// TIA Portal V20 export
FUNCTION_BLOCK "PR_LoadingSeq_Soft2.0 1_workflow_95d36b"   // FB48, LAD
{ S7_Optimized_Access := 'TRUE' }
// stored: MemoryReserve 100, SetENOAutomatically false
   VAR_INPUT
      iAbort : Bool;
      iAcceptPartPresent : Bool;
      iAutoRunning : Bool;
      iFaultReset : Bool;
      iLoadGantrySafe : Bool;
      iOTS_Frm_Prev : Bool;
      iPartPresent : Bool;
      iPartPresentInGrip : Bool;
      iRFWriteDone : Bool;
      iRFWriteError : Bool;
      iReject : Bool;
      iReset_fault : Bool;
      iRetry : Bool;
      iRetryCount : Int;
      iSstMode : Bool;
      iSstPB : Bool;
      iStartFrmFibroseq : Bool;
   END_VAR
   VAR_OUTPUT
      qError : Array[0..1] of Bool;
      qLoadingOver : Bool;
      qMessage : Array[0..1] of Bool;
      qRTR_To_Prev : Bool;
   END_VAR
   VAR
      c121_WaitForRFIDWriteOver_T1 : Bool;
      c121_WaitForRFIDWriteOver_T2 : Bool;
      c122_CheckRetryCountOver_T1 : Bool;
      c122_CheckRetryCountOver_T2 : Bool;
      c123_WaitForOperatorDecision_T1 : Bool;
      c123_WaitForOperatorDecision_T2 : Bool;
      c20_CheckRecoveryStatus_T1 : Bool;
      c20_CheckRecoveryStatus_T2 : Bool;
      c20_CheckRecoveryStatus_T3 : Bool;
      c50_CheckPartPresentAtStation_T1 : Bool;
      c50_CheckPartPresentAtStation_T2 : Bool;
      c90_ConfirmPartLoad_T1 : Bool;
      c90_ConfirmPartLoad_T2 : Bool;
      StateNo : Int;
      s100_WaitForOperatorDecision : Bool;
      s100_WaitForOperatorDecision_T1 : Bool;
      s100_WaitForOperatorDecision_T2 : Bool;
      s10_WaitForStartFrmFibroMainSeq : Bool;
      s10_WaitForStartFrmFibroMainSeq_T1 : Bool;
      s120_WaitForGantrySafe : Bool;
      s120_WaitForGantrySafe_T1 : Bool;
      s121_WaitForRFIDWriteOver : Bool;
      s121_WaitForRFIDWriteOver_T1 : Bool;
      s121_WaitForRFIDWriteOver_T2 : Bool;
      s122_CheckRetryCountOver : Bool;
      s122_CheckRetryCountOver_T1 : Bool;
      s122_CheckRetryCountOver_T2 : Bool;
      s123_WaitForOperatorDecision : Bool;
      s123_WaitForOperatorDecision_T1 : Bool;
      s123_WaitForOperatorDecision_T2 : Bool;
      s130_WaitForStartLow : Bool;
      s130_WaitForStartLow_T1 : Bool;
      s1_WaitForResetRelease : Bool;
      s1_WaitForResetRelease_T1 : Bool;
      s20_CheckRecoveryStatus : Bool;
      s20_CheckRecoveryStatus_T1 : Bool;
      s20_CheckRecoveryStatus_T2 : Bool;
      s20_CheckRecoveryStatus_T3 : Bool;
      s30_WaitForOperatorAck : Bool;
      s30_WaitForOperatorAck_T1 : Bool;
      s40_WaitForLoadingGantrySafe : Bool;
      s40_WaitForLoadingGantrySafe_T1 : Bool;
      s50_CheckPartPresentAtStation : Bool;
      s50_CheckPartPresentAtStation_T1 : Bool;
      s50_CheckPartPresentAtStation_T2 : Bool;
      s60_WaitForPartAbsentAndAck : Bool;
      s60_WaitForPartAbsentAndAck_T1 : Bool;
      s70_WaitForOTSFromGantry : Bool;
      s70_WaitForOTSFromGantry_T1 : Bool;
      s80_WaitForPartLoad : Bool;
      s80_WaitForPartLoad_T1 : Bool;
      s90_ConfirmPartLoad : Bool;
      s90_ConfirmPartLoad_T1 : Bool;
      s90_ConfirmPartLoad_T2 : Bool;
      sAbnormalStatus : Bool;
      sLoadInProgress : Bool;
      sLoadInProgressInternal : Int;
      sPartPresent : Bool;
      sRFWriteRetryCount : Int;
      sSst : Bool;
      sSstPulse : Bool;
      sSstRise : Bool;
      sStWtResetRel : Bool;
      sStWtResetRel_T1 : Bool;
   END_VAR
   VAR_TEMP
      tOne : Bool;
   END_VAR
   VAR_TEMP   // added for the SCL form of the ladder/FBD networks
      _w1 : Bool;
      _w2 : Bool;
   END_VAR
BEGIN

REGION Network 1
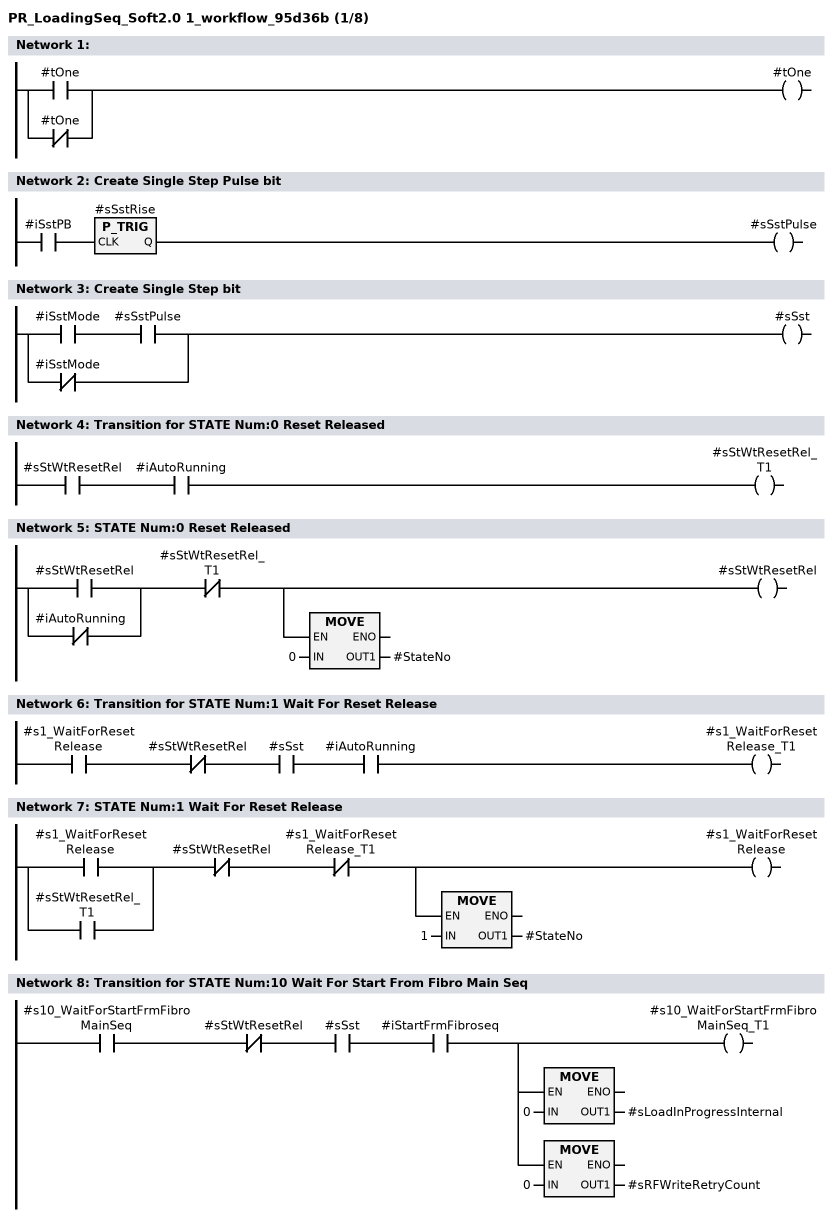
   RUNG wire#powerrail
      Contact( #tOne )
      wire#w1
      Coil( #tOne )
   END_RUNG
   RUNG wire#powerrail
      I_Contact( #tOne )
   END_RUNG wire#w1
   // the same network as SCL:
   #tOne := #tOne OR NOT #tOne;
END_REGION

REGION Network 2: Create Single Step Pulse bit
   RUNG wire#powerrail
      Contact( #iSstPB )
      P_Trig( #sSstRise )
      Coil( #sSstPulse )
   END_RUNG
   // the same network as SCL:
   #_w1 := #iSstPB AND NOT #sSstRise;   // rising edge
   #sSstRise := #iSstPB;
   #sSstPulse := #_w1;
END_REGION

REGION Network 3: Create Single Step bit
   RUNG wire#powerrail
      Contact( #iSstMode )
      Contact( #sSstPulse )
      wire#w1
      Coil( #sSst )
   END_RUNG
   RUNG wire#powerrail
      I_Contact( #iSstMode )
   END_RUNG wire#w1
   // the same network as SCL:
   #sSst := (#iSstMode AND #sSstPulse) OR NOT #iSstMode;
END_REGION

REGION Network 4: Transition for STATE Num:0 Reset Released
   RUNG wire#powerrail
      Contact( #sStWtResetRel )
      Contact( #iAutoRunning )
      Coil( #sStWtResetRel_T1 )
   END_RUNG
   // the same network as SCL:
   #sStWtResetRel_T1 := #sStWtResetRel AND #iAutoRunning;
END_REGION

REGION Network 5: STATE Num:0 Reset Released
   RUNG wire#powerrail
      Contact( #sStWtResetRel )
      wire#w1
      I_Contact( #sStWtResetRel_T1 )
      wire#w2
      Coil( #sStWtResetRel )
   END_RUNG
   RUNG wire#powerrail
      I_Contact( #iAutoRunning )
   END_RUNG wire#w1
   RUNG wire#w2
      { S7_GenerateENO := "TRUE" } Move(in := 0, out1 => #StateNo)
   END_RUNG
   // the same network as SCL:
   #sStWtResetRel := (#sStWtResetRel OR NOT #iAutoRunning) AND NOT #sStWtResetRel_T1;
   IF #sStWtResetRel THEN #StateNo := 0; END_IF;
END_REGION

REGION Network 6: Transition for STATE Num:1 Wait For Reset Release
   RUNG wire#powerrail
      Contact( #s1_WaitForResetRelease )
      I_Contact( #sStWtResetRel )
      Contact( #sSst )
      Contact( #iAutoRunning )
      Coil( #s1_WaitForResetRelease_T1 )
   END_RUNG
   // the same network as SCL:
   #s1_WaitForResetRelease_T1 := #s1_WaitForResetRelease AND NOT #sStWtResetRel AND #sSst AND #iAutoRunning;
END_REGION

REGION Network 7: STATE Num:1 Wait For Reset Release
   RUNG wire#powerrail
      Contact( #s1_WaitForResetRelease )
      wire#w1
      I_Contact( #sStWtResetRel )
      I_Contact( #s1_WaitForResetRelease_T1 )
      wire#w2
      Coil( #s1_WaitForResetRelease )
   END_RUNG
   RUNG wire#powerrail
      Contact( #sStWtResetRel_T1 )
   END_RUNG wire#w1
   RUNG wire#w2
      { S7_GenerateENO := "TRUE" } Move(in := 1, out1 => #StateNo)
   END_RUNG
   // the same network as SCL:
   #s1_WaitForResetRelease := (#s1_WaitForResetRelease OR #sStWtResetRel_T1) AND NOT #sStWtResetRel AND NOT #s1_WaitForResetRelease_T1;
   IF #s1_WaitForResetRelease THEN #StateNo := 1; END_IF;
END_REGION

REGION Network 8: Transition for STATE Num:10 Wait For Start From Fibro Main Seq
   RUNG wire#powerrail
      Contact( #s10_WaitForStartFrmFibroMainSeq )
      I_Contact( #sStWtResetRel )
      Contact( #sSst )
      Contact( #iStartFrmFibroseq )
      wire#w1
      Coil( #s10_WaitForStartFrmFibroMainSeq_T1 )
   END_RUNG
   RUNG wire#w1
      Move(in := 0, out1 => #sLoadInProgressInternal)
   END_RUNG
   RUNG wire#w1
      Move(in := 0, out1 => #sRFWriteRetryCount)
   END_RUNG
   // the same network as SCL:
   #s10_WaitForStartFrmFibroMainSeq_T1 := #s10_WaitForStartFrmFibroMainSeq AND NOT #sStWtResetRel AND #sSst AND #iStartFrmFibroseq;
   IF #s10_WaitForStartFrmFibroMainSeq_T1 THEN
       #sLoadInProgressInternal := 0;
       #sRFWriteRetryCount := 0;
   END_IF;
END_REGION

REGION Network 9: STATE Num:10 Wait For Start From Fibro Main Seq
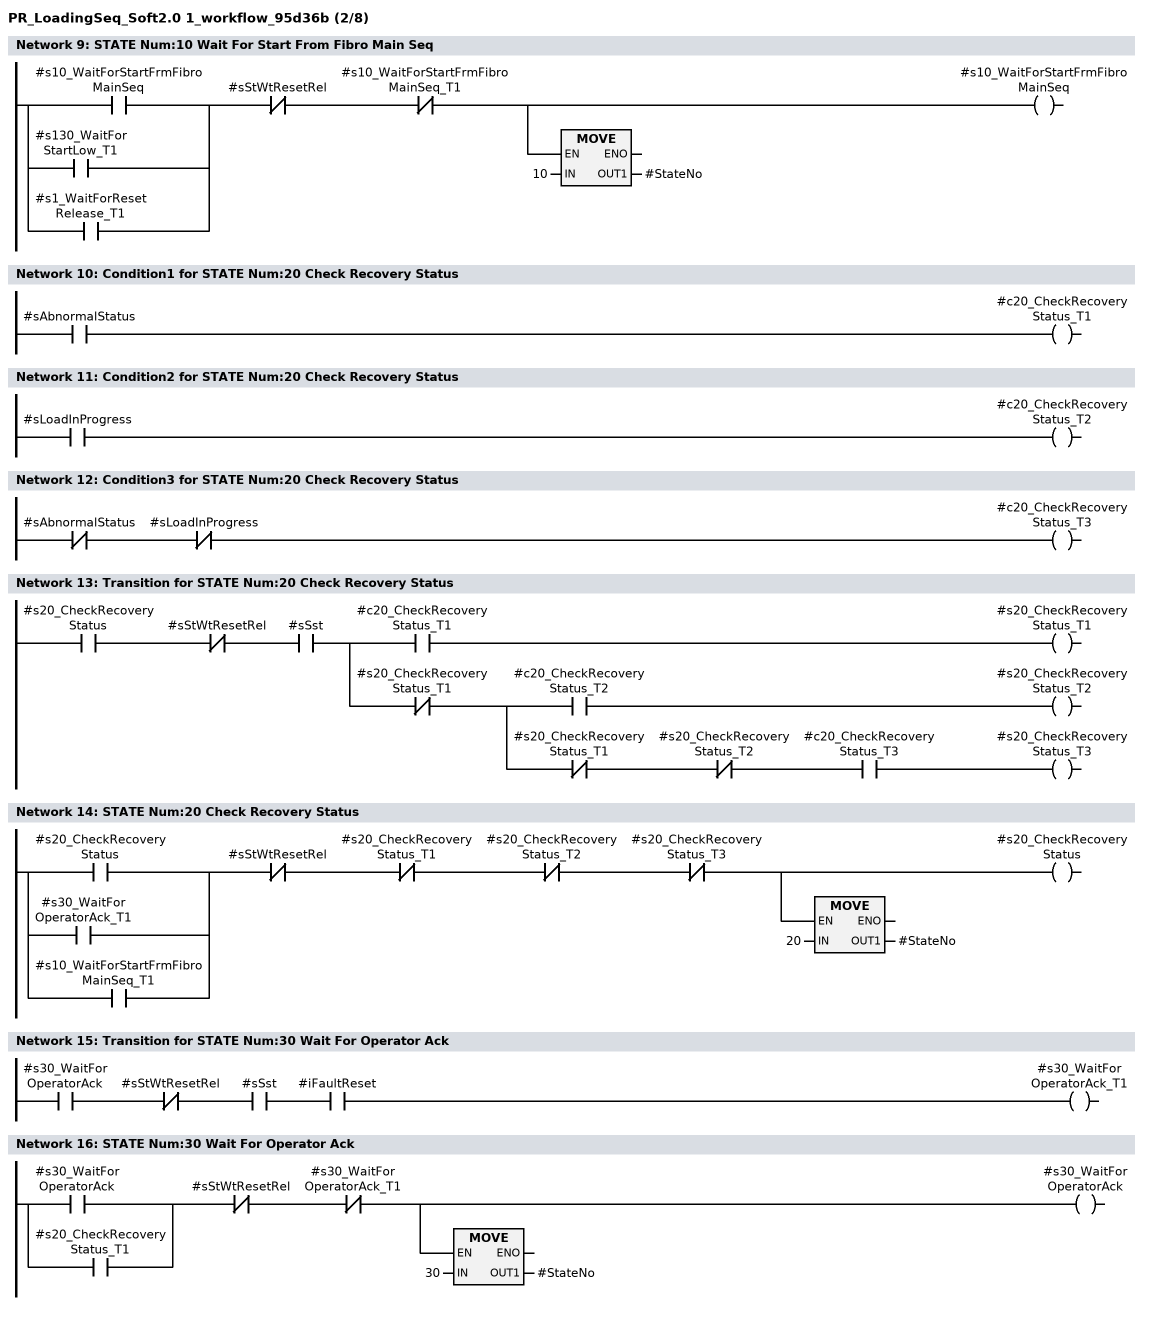
   RUNG wire#powerrail
      Contact( #s10_WaitForStartFrmFibroMainSeq )
      wire#w1
      I_Contact( #sStWtResetRel )
      I_Contact( #s10_WaitForStartFrmFibroMainSeq_T1 )
      wire#w2
      Coil( #s10_WaitForStartFrmFibroMainSeq )
   END_RUNG
   RUNG wire#powerrail
      Contact( #s130_WaitForStartLow_T1 )
   END_RUNG wire#w1
   RUNG wire#powerrail
      Contact( #s1_WaitForResetRelease_T1 )
   END_RUNG wire#w1
   RUNG wire#w2
      { S7_GenerateENO := "TRUE" } Move(in := 10, out1 => #StateNo)
   END_RUNG
   // the same network as SCL:
   #s10_WaitForStartFrmFibroMainSeq := (#s10_WaitForStartFrmFibroMainSeq OR #s130_WaitForStartLow_T1 OR #s1_WaitForResetRelease_T1) AND NOT #sStWtResetRel AND NOT #s10_WaitForStartFrmFibroMainSeq_T1;
   IF #s10_WaitForStartFrmFibroMainSeq THEN #StateNo := 10; END_IF;
END_REGION

REGION Network 10: Condition1 for STATE Num:20 Check Recovery Status
   RUNG wire#powerrail
      Contact( #sAbnormalStatus )
      Coil( #c20_CheckRecoveryStatus_T1 )
   END_RUNG
   // the same network as SCL:
   #c20_CheckRecoveryStatus_T1 := #sAbnormalStatus;
END_REGION

REGION Network 11: Condition2 for STATE Num:20 Check Recovery Status
   RUNG wire#powerrail
      Contact( #sLoadInProgress )
      Coil( #c20_CheckRecoveryStatus_T2 )
   END_RUNG
   // the same network as SCL:
   #c20_CheckRecoveryStatus_T2 := #sLoadInProgress;
END_REGION

REGION Network 12: Condition3 for STATE Num:20 Check Recovery Status
   RUNG wire#powerrail
      I_Contact( #sAbnormalStatus )
      I_Contact( #sLoadInProgress )
      Coil( #c20_CheckRecoveryStatus_T3 )
   END_RUNG
   // the same network as SCL:
   #c20_CheckRecoveryStatus_T3 := NOT #sAbnormalStatus AND NOT #sLoadInProgress;
END_REGION

REGION Network 13: Transition for STATE Num:20 Check Recovery Status
   RUNG wire#powerrail
      Contact( #s20_CheckRecoveryStatus )
      I_Contact( #sStWtResetRel )
      Contact( #sSst )
      wire#w1
      Contact( #c20_CheckRecoveryStatus_T1 )
      Coil( #s20_CheckRecoveryStatus_T1 )
   END_RUNG
   RUNG wire#w1
      I_Contact( #s20_CheckRecoveryStatus_T1 )
      wire#w2
      Contact( #c20_CheckRecoveryStatus_T2 )
      Coil( #s20_CheckRecoveryStatus_T2 )
   END_RUNG
   RUNG wire#w2
      I_Contact( #s20_CheckRecoveryStatus_T1 )
      I_Contact( #s20_CheckRecoveryStatus_T2 )
      Contact( #c20_CheckRecoveryStatus_T3 )
      Coil( #s20_CheckRecoveryStatus_T3 )
   END_RUNG
   // the same network as SCL:
   #_w1 := #s20_CheckRecoveryStatus AND NOT #sStWtResetRel AND #sSst;
   #s20_CheckRecoveryStatus_T1 := #_w1 AND #c20_CheckRecoveryStatus_T1;
   #_w2 := #_w1 AND NOT #s20_CheckRecoveryStatus_T1;
   #s20_CheckRecoveryStatus_T2 := #_w2 AND #c20_CheckRecoveryStatus_T2;
   #s20_CheckRecoveryStatus_T3 := #_w2 AND NOT #s20_CheckRecoveryStatus_T1 AND NOT #s20_CheckRecoveryStatus_T2 AND #c20_CheckRecoveryStatus_T3;
END_REGION

REGION Network 14: STATE Num:20 Check Recovery Status
   RUNG wire#powerrail
      Contact( #s20_CheckRecoveryStatus )
      wire#w1
      I_Contact( #sStWtResetRel )
      I_Contact( #s20_CheckRecoveryStatus_T1 )
      I_Contact( #s20_CheckRecoveryStatus_T2 )
      I_Contact( #s20_CheckRecoveryStatus_T3 )
      wire#w2
      Coil( #s20_CheckRecoveryStatus )
   END_RUNG
   RUNG wire#powerrail
      Contact( #s30_WaitForOperatorAck_T1 )
   END_RUNG wire#w1
   RUNG wire#powerrail
      Contact( #s10_WaitForStartFrmFibroMainSeq_T1 )
   END_RUNG wire#w1
   RUNG wire#w2
      { S7_GenerateENO := "TRUE" } Move(in := 20, out1 => #StateNo)
   END_RUNG
   // the same network as SCL:
   #s20_CheckRecoveryStatus := (#s20_CheckRecoveryStatus OR #s30_WaitForOperatorAck_T1 OR #s10_WaitForStartFrmFibroMainSeq_T1) AND NOT #sStWtResetRel AND NOT #s20_CheckRecoveryStatus_T1 AND NOT #s20_CheckRecoveryStatus_T2 AND NOT #s20_CheckRecoveryStatus_T3;
   IF #s20_CheckRecoveryStatus THEN #StateNo := 20; END_IF;
END_REGION

REGION Network 15: Transition for STATE Num:30 Wait For Operator Ack
   RUNG wire#powerrail
      Contact( #s30_WaitForOperatorAck )
      I_Contact( #sStWtResetRel )
      Contact( #sSst )
      Contact( #iFaultReset )
      Coil( #s30_WaitForOperatorAck_T1 )
   END_RUNG
   // the same network as SCL:
   #s30_WaitForOperatorAck_T1 := #s30_WaitForOperatorAck AND NOT #sStWtResetRel AND #sSst AND #iFaultReset;
END_REGION

REGION Network 16: STATE Num:30 Wait For Operator Ack
   RUNG wire#powerrail
      Contact( #s30_WaitForOperatorAck )
      wire#w1
      I_Contact( #sStWtResetRel )
      I_Contact( #s30_WaitForOperatorAck_T1 )
      wire#w2
      Coil( #s30_WaitForOperatorAck )
   END_RUNG
   RUNG wire#powerrail
      Contact( #s20_CheckRecoveryStatus_T1 )
   END_RUNG wire#w1
   RUNG wire#w2
      { S7_GenerateENO := "TRUE" } Move(in := 30, out1 => #StateNo)
   END_RUNG
   // the same network as SCL:
   #s30_WaitForOperatorAck := (#s30_WaitForOperatorAck OR #s20_CheckRecoveryStatus_T1) AND NOT #sStWtResetRel AND NOT #s30_WaitForOperatorAck_T1;
   IF #s30_WaitForOperatorAck THEN #StateNo := 30; END_IF;
END_REGION

REGION Network 17: Actions for STATE Num:30 Wait For Operator Ack
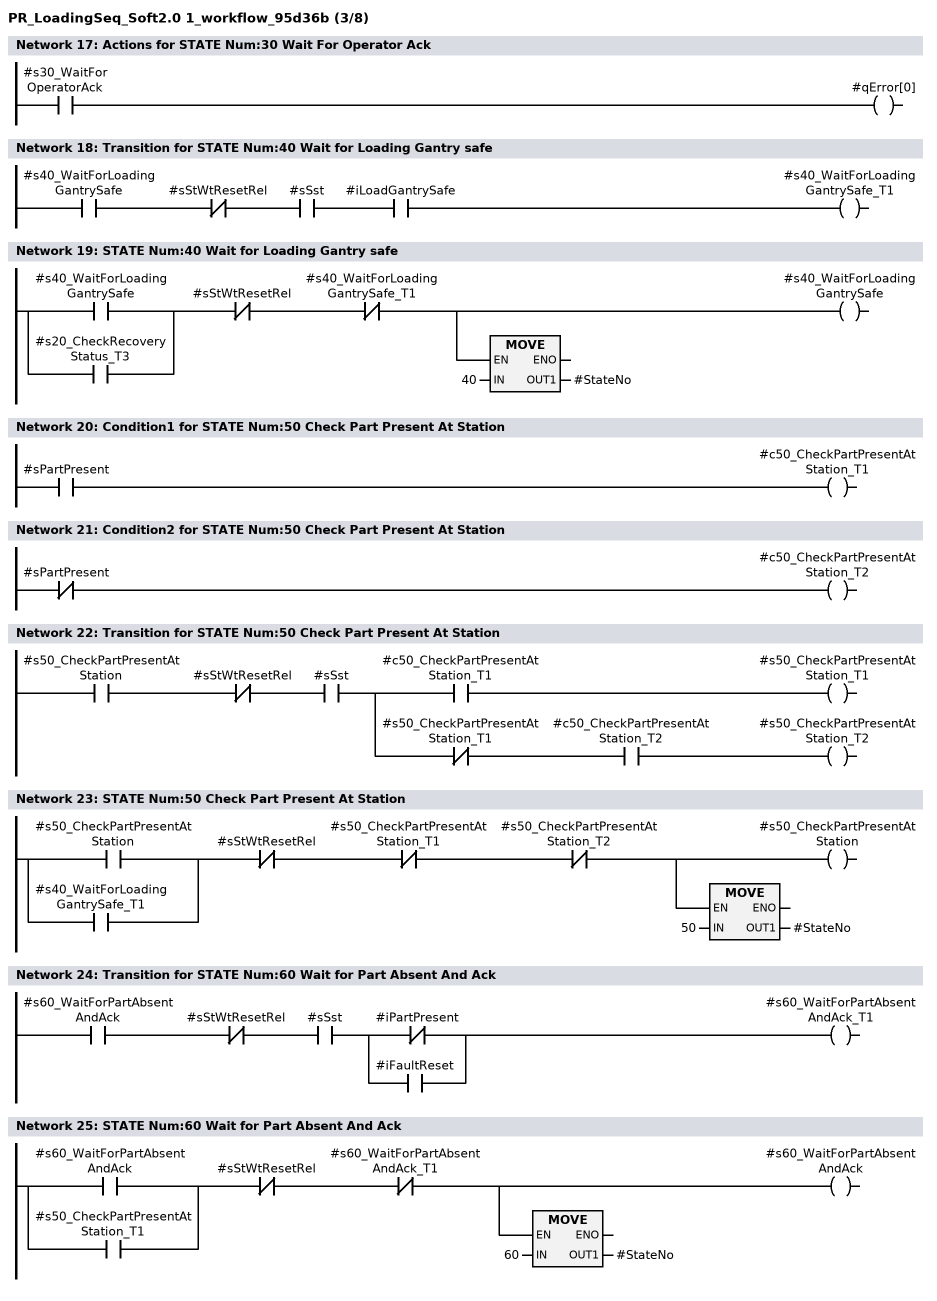
   RUNG wire#powerrail
      Contact( #s30_WaitForOperatorAck )
      Coil( #qError[0] )
   END_RUNG
   // the same network as SCL:
   #qError[0] := #s30_WaitForOperatorAck;
END_REGION

REGION Network 18: Transition for STATE Num:40 Wait for Loading Gantry safe
   RUNG wire#powerrail
      Contact( #s40_WaitForLoadingGantrySafe )
      I_Contact( #sStWtResetRel )
      Contact( #sSst )
      Contact( #iLoadGantrySafe )
      Coil( #s40_WaitForLoadingGantrySafe_T1 )
   END_RUNG
   // the same network as SCL:
   #s40_WaitForLoadingGantrySafe_T1 := #s40_WaitForLoadingGantrySafe AND NOT #sStWtResetRel AND #sSst AND #iLoadGantrySafe;
END_REGION

REGION Network 19: STATE Num:40 Wait for Loading Gantry safe
   RUNG wire#powerrail
      Contact( #s40_WaitForLoadingGantrySafe )
      wire#w1
      I_Contact( #sStWtResetRel )
      I_Contact( #s40_WaitForLoadingGantrySafe_T1 )
      wire#w2
      Coil( #s40_WaitForLoadingGantrySafe )
   END_RUNG
   RUNG wire#powerrail
      Contact( #s20_CheckRecoveryStatus_T3 )
   END_RUNG wire#w1
   RUNG wire#w2
      { S7_GenerateENO := "TRUE" } Move(in := 40, out1 => #StateNo)
   END_RUNG
   // the same network as SCL:
   #s40_WaitForLoadingGantrySafe := (#s40_WaitForLoadingGantrySafe OR #s20_CheckRecoveryStatus_T3) AND NOT #sStWtResetRel AND NOT #s40_WaitForLoadingGantrySafe_T1;
   IF #s40_WaitForLoadingGantrySafe THEN #StateNo := 40; END_IF;
END_REGION

REGION Network 20: Condition1 for STATE Num:50 Check Part Present At Station
   RUNG wire#powerrail
      Contact( #sPartPresent )
      Coil( #c50_CheckPartPresentAtStation_T1 )
   END_RUNG
   // the same network as SCL:
   #c50_CheckPartPresentAtStation_T1 := #sPartPresent;
END_REGION

REGION Network 21: Condition2 for STATE Num:50 Check Part Present At Station
   RUNG wire#powerrail
      I_Contact( #sPartPresent )
      Coil( #c50_CheckPartPresentAtStation_T2 )
   END_RUNG
   // the same network as SCL:
   #c50_CheckPartPresentAtStation_T2 := NOT #sPartPresent;
END_REGION

REGION Network 22: Transition for STATE Num:50 Check Part Present At Station
   RUNG wire#powerrail
      Contact( #s50_CheckPartPresentAtStation )
      I_Contact( #sStWtResetRel )
      Contact( #sSst )
      wire#w1
      Contact( #c50_CheckPartPresentAtStation_T1 )
      Coil( #s50_CheckPartPresentAtStation_T1 )
   END_RUNG
   RUNG wire#w1
      I_Contact( #s50_CheckPartPresentAtStation_T1 )
      Contact( #c50_CheckPartPresentAtStation_T2 )
      Coil( #s50_CheckPartPresentAtStation_T2 )
   END_RUNG
   // the same network as SCL:
   #_w1 := #s50_CheckPartPresentAtStation AND NOT #sStWtResetRel AND #sSst;
   #s50_CheckPartPresentAtStation_T1 := #_w1 AND #c50_CheckPartPresentAtStation_T1;
   #s50_CheckPartPresentAtStation_T2 := #_w1 AND NOT #s50_CheckPartPresentAtStation_T1 AND #c50_CheckPartPresentAtStation_T2;
END_REGION

REGION Network 23: STATE Num:50 Check Part Present At Station
   RUNG wire#powerrail
      Contact( #s50_CheckPartPresentAtStation )
      wire#w1
      I_Contact( #sStWtResetRel )
      I_Contact( #s50_CheckPartPresentAtStation_T1 )
      I_Contact( #s50_CheckPartPresentAtStation_T2 )
      wire#w2
      Coil( #s50_CheckPartPresentAtStation )
   END_RUNG
   RUNG wire#powerrail
      Contact( #s40_WaitForLoadingGantrySafe_T1 )
   END_RUNG wire#w1
   RUNG wire#w2
      { S7_GenerateENO := "TRUE" } Move(in := 50, out1 => #StateNo)
   END_RUNG
   // the same network as SCL:
   #s50_CheckPartPresentAtStation := (#s50_CheckPartPresentAtStation OR #s40_WaitForLoadingGantrySafe_T1) AND NOT #sStWtResetRel AND NOT #s50_CheckPartPresentAtStation_T1 AND NOT #s50_CheckPartPresentAtStation_T2;
   IF #s50_CheckPartPresentAtStation THEN #StateNo := 50; END_IF;
END_REGION

REGION Network 24: Transition for STATE Num:60 Wait for Part Absent And Ack
   RUNG wire#powerrail
      Contact( #s60_WaitForPartAbsentAndAck )
      I_Contact( #sStWtResetRel )
      Contact( #sSst )
      wire#w1
      I_Contact( #iPartPresent )
      wire#w2
      Coil( #s60_WaitForPartAbsentAndAck_T1 )
   END_RUNG
   RUNG wire#w1
      Contact( #iFaultReset )
   END_RUNG wire#w2
   // the same network as SCL:
   #s60_WaitForPartAbsentAndAck_T1 := #s60_WaitForPartAbsentAndAck AND NOT #sStWtResetRel AND #sSst AND (NOT #iPartPresent OR #iFaultReset);
END_REGION

REGION Network 25: STATE Num:60 Wait for Part Absent And Ack
   RUNG wire#powerrail
      Contact( #s60_WaitForPartAbsentAndAck )
      wire#w1
      I_Contact( #sStWtResetRel )
      I_Contact( #s60_WaitForPartAbsentAndAck_T1 )
      wire#w2
      Coil( #s60_WaitForPartAbsentAndAck )
   END_RUNG
   RUNG wire#powerrail
      Contact( #s50_CheckPartPresentAtStation_T1 )
   END_RUNG wire#w1
   RUNG wire#w2
      { S7_GenerateENO := "TRUE" } Move(in := 60, out1 => #StateNo)
   END_RUNG
   // the same network as SCL:
   #s60_WaitForPartAbsentAndAck := (#s60_WaitForPartAbsentAndAck OR #s50_CheckPartPresentAtStation_T1) AND NOT #sStWtResetRel AND NOT #s60_WaitForPartAbsentAndAck_T1;
   IF #s60_WaitForPartAbsentAndAck THEN #StateNo := 60; END_IF;
END_REGION

REGION Network 26: Transition for STATE Num:70 Wait For OTS From Gantry
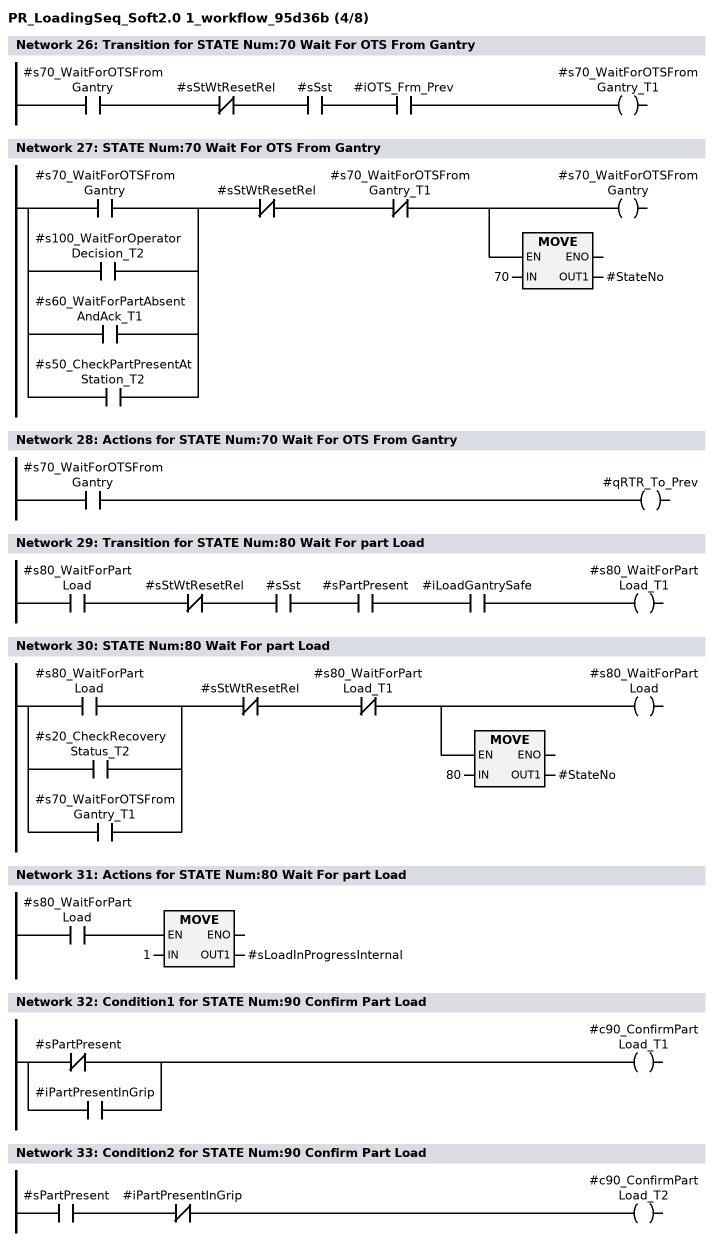
   RUNG wire#powerrail
      Contact( #s70_WaitForOTSFromGantry )
      I_Contact( #sStWtResetRel )
      Contact( #sSst )
      Contact( #iOTS_Frm_Prev )
      Coil( #s70_WaitForOTSFromGantry_T1 )
   END_RUNG
   // the same network as SCL:
   #s70_WaitForOTSFromGantry_T1 := #s70_WaitForOTSFromGantry AND NOT #sStWtResetRel AND #sSst AND #iOTS_Frm_Prev;
END_REGION

REGION Network 27: STATE Num:70 Wait For OTS From Gantry
   RUNG wire#powerrail
      Contact( #s70_WaitForOTSFromGantry )
      wire#w1
      I_Contact( #sStWtResetRel )
      I_Contact( #s70_WaitForOTSFromGantry_T1 )
      wire#w2
      Coil( #s70_WaitForOTSFromGantry )
   END_RUNG
   RUNG wire#powerrail
      Contact( #s100_WaitForOperatorDecision_T2 )
   END_RUNG wire#w1
   RUNG wire#powerrail
      Contact( #s60_WaitForPartAbsentAndAck_T1 )
   END_RUNG wire#w1
   RUNG wire#powerrail
      Contact( #s50_CheckPartPresentAtStation_T2 )
   END_RUNG wire#w1
   RUNG wire#w2
      { S7_GenerateENO := "TRUE" } Move(in := 70, out1 => #StateNo)
   END_RUNG
   // the same network as SCL:
   #s70_WaitForOTSFromGantry := (#s70_WaitForOTSFromGantry OR #s100_WaitForOperatorDecision_T2 OR #s60_WaitForPartAbsentAndAck_T1 OR #s50_CheckPartPresentAtStation_T2) AND NOT #sStWtResetRel AND NOT #s70_WaitForOTSFromGantry_T1;
   IF #s70_WaitForOTSFromGantry THEN #StateNo := 70; END_IF;
END_REGION

REGION Network 28: Actions for STATE Num:70 Wait For OTS From Gantry
   RUNG wire#powerrail
      Contact( #s70_WaitForOTSFromGantry )
      Coil( #qRTR_To_Prev )
   END_RUNG
   // the same network as SCL:
   #qRTR_To_Prev := #s70_WaitForOTSFromGantry;
END_REGION

REGION Network 29: Transition for STATE Num:80 Wait For part Load
   RUNG wire#powerrail
      Contact( #s80_WaitForPartLoad )
      I_Contact( #sStWtResetRel )
      Contact( #sSst )
      Contact( #sPartPresent )
      Contact( #iLoadGantrySafe )
      Coil( #s80_WaitForPartLoad_T1 )
   END_RUNG
   // the same network as SCL:
   #s80_WaitForPartLoad_T1 := #s80_WaitForPartLoad AND NOT #sStWtResetRel AND #sSst AND #sPartPresent AND #iLoadGantrySafe;
END_REGION

REGION Network 30: STATE Num:80 Wait For part Load
   RUNG wire#powerrail
      Contact( #s80_WaitForPartLoad )
      wire#w1
      I_Contact( #sStWtResetRel )
      I_Contact( #s80_WaitForPartLoad_T1 )
      wire#w2
      Coil( #s80_WaitForPartLoad )
   END_RUNG
   RUNG wire#powerrail
      Contact( #s20_CheckRecoveryStatus_T2 )
   END_RUNG wire#w1
   RUNG wire#powerrail
      Contact( #s70_WaitForOTSFromGantry_T1 )
   END_RUNG wire#w1
   RUNG wire#w2
      { S7_GenerateENO := "TRUE" } Move(in := 80, out1 => #StateNo)
   END_RUNG
   // the same network as SCL:
   #s80_WaitForPartLoad := (#s80_WaitForPartLoad OR #s20_CheckRecoveryStatus_T2 OR #s70_WaitForOTSFromGantry_T1) AND NOT #sStWtResetRel AND NOT #s80_WaitForPartLoad_T1;
   IF #s80_WaitForPartLoad THEN #StateNo := 80; END_IF;
END_REGION

REGION Network 31: Actions for STATE Num:80 Wait For part Load
   RUNG wire#powerrail
      Contact( #s80_WaitForPartLoad )
      { S7_GenerateENO := "TRUE" } Move(in := 1, out1 => #sLoadInProgressInternal)
   END_RUNG
   // the same network as SCL:
   IF #s80_WaitForPartLoad THEN #sLoadInProgressInternal := 1; END_IF;
END_REGION

REGION Network 32: Condition1 for STATE Num:90 Confirm Part Load
   RUNG wire#powerrail
      I_Contact( #sPartPresent )
      wire#w1
      Coil( #c90_ConfirmPartLoad_T1 )
   END_RUNG
   RUNG wire#powerrail
      Contact( #iPartPresentInGrip )
   END_RUNG wire#w1
   // the same network as SCL:
   #c90_ConfirmPartLoad_T1 := NOT #sPartPresent OR #iPartPresentInGrip;
END_REGION

REGION Network 33: Condition2 for STATE Num:90 Confirm Part Load
   RUNG wire#powerrail
      Contact( #sPartPresent )
      I_Contact( #iPartPresentInGrip )
      Coil( #c90_ConfirmPartLoad_T2 )
   END_RUNG
   // the same network as SCL:
   #c90_ConfirmPartLoad_T2 := #sPartPresent AND NOT #iPartPresentInGrip;
END_REGION

REGION Network 34: Transition for STATE Num:90 Confirm Part Load
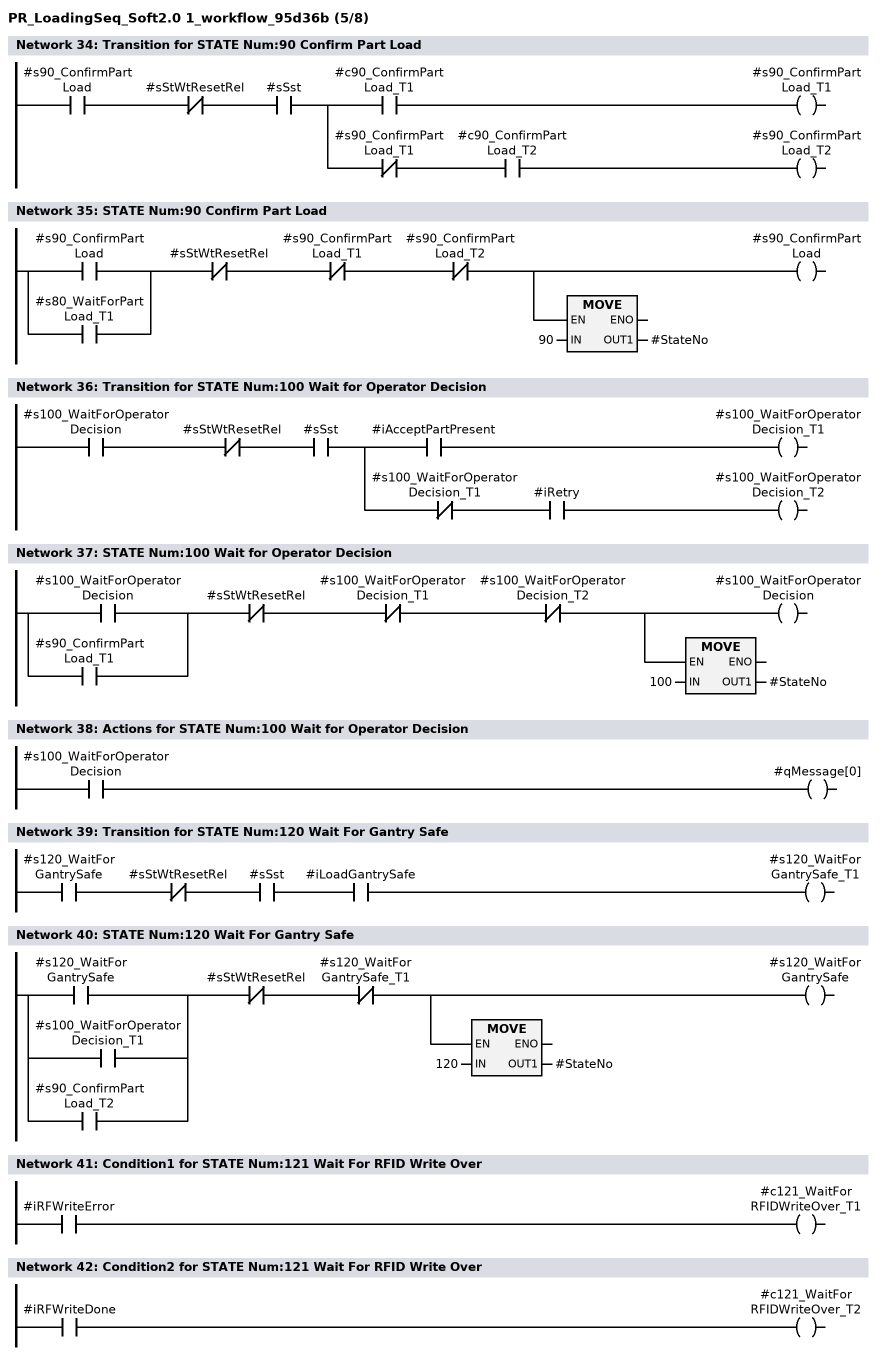
   RUNG wire#powerrail
      Contact( #s90_ConfirmPartLoad )
      I_Contact( #sStWtResetRel )
      Contact( #sSst )
      wire#w1
      Contact( #c90_ConfirmPartLoad_T1 )
      Coil( #s90_ConfirmPartLoad_T1 )
   END_RUNG
   RUNG wire#w1
      I_Contact( #s90_ConfirmPartLoad_T1 )
      Contact( #c90_ConfirmPartLoad_T2 )
      Coil( #s90_ConfirmPartLoad_T2 )
   END_RUNG
   // the same network as SCL:
   #_w1 := #s90_ConfirmPartLoad AND NOT #sStWtResetRel AND #sSst;
   #s90_ConfirmPartLoad_T1 := #_w1 AND #c90_ConfirmPartLoad_T1;
   #s90_ConfirmPartLoad_T2 := #_w1 AND NOT #s90_ConfirmPartLoad_T1 AND #c90_ConfirmPartLoad_T2;
END_REGION

REGION Network 35: STATE Num:90 Confirm Part Load
   RUNG wire#powerrail
      Contact( #s90_ConfirmPartLoad )
      wire#w1
      I_Contact( #sStWtResetRel )
      I_Contact( #s90_ConfirmPartLoad_T1 )
      I_Contact( #s90_ConfirmPartLoad_T2 )
      wire#w2
      Coil( #s90_ConfirmPartLoad )
   END_RUNG
   RUNG wire#powerrail
      Contact( #s80_WaitForPartLoad_T1 )
   END_RUNG wire#w1
   RUNG wire#w2
      { S7_GenerateENO := "TRUE" } Move(in := 90, out1 => #StateNo)
   END_RUNG
   // the same network as SCL:
   #s90_ConfirmPartLoad := (#s90_ConfirmPartLoad OR #s80_WaitForPartLoad_T1) AND NOT #sStWtResetRel AND NOT #s90_ConfirmPartLoad_T1 AND NOT #s90_ConfirmPartLoad_T2;
   IF #s90_ConfirmPartLoad THEN #StateNo := 90; END_IF;
END_REGION

REGION Network 36: Transition for STATE Num:100 Wait for Operator Decision
   RUNG wire#powerrail
      Contact( #s100_WaitForOperatorDecision )
      I_Contact( #sStWtResetRel )
      Contact( #sSst )
      wire#w1
      Contact( #iAcceptPartPresent )
      Coil( #s100_WaitForOperatorDecision_T1 )
   END_RUNG
   RUNG wire#w1
      I_Contact( #s100_WaitForOperatorDecision_T1 )
      Contact( #iRetry )
      Coil( #s100_WaitForOperatorDecision_T2 )
   END_RUNG
   // the same network as SCL:
   #_w1 := #s100_WaitForOperatorDecision AND NOT #sStWtResetRel AND #sSst;
   #s100_WaitForOperatorDecision_T1 := #_w1 AND #iAcceptPartPresent;
   #s100_WaitForOperatorDecision_T2 := #_w1 AND NOT #s100_WaitForOperatorDecision_T1 AND #iRetry;
END_REGION

REGION Network 37: STATE Num:100 Wait for Operator Decision
   RUNG wire#powerrail
      Contact( #s100_WaitForOperatorDecision )
      wire#w1
      I_Contact( #sStWtResetRel )
      I_Contact( #s100_WaitForOperatorDecision_T1 )
      I_Contact( #s100_WaitForOperatorDecision_T2 )
      wire#w2
      Coil( #s100_WaitForOperatorDecision )
   END_RUNG
   RUNG wire#powerrail
      Contact( #s90_ConfirmPartLoad_T1 )
   END_RUNG wire#w1
   RUNG wire#w2
      { S7_GenerateENO := "TRUE" } Move(in := 100, out1 => #StateNo)
   END_RUNG
   // the same network as SCL:
   #s100_WaitForOperatorDecision := (#s100_WaitForOperatorDecision OR #s90_ConfirmPartLoad_T1) AND NOT #sStWtResetRel AND NOT #s100_WaitForOperatorDecision_T1 AND NOT #s100_WaitForOperatorDecision_T2;
   IF #s100_WaitForOperatorDecision THEN #StateNo := 100; END_IF;
END_REGION

REGION Network 38: Actions for STATE Num:100 Wait for Operator Decision
   RUNG wire#powerrail
      Contact( #s100_WaitForOperatorDecision )
      Coil( #qMessage[0] )
   END_RUNG
   // the same network as SCL:
   #qMessage[0] := #s100_WaitForOperatorDecision;
END_REGION

REGION Network 39: Transition for STATE Num:120 Wait For Gantry Safe
   RUNG wire#powerrail
      Contact( #s120_WaitForGantrySafe )
      I_Contact( #sStWtResetRel )
      Contact( #sSst )
      Contact( #iLoadGantrySafe )
      Coil( #s120_WaitForGantrySafe_T1 )
   END_RUNG
   // the same network as SCL:
   #s120_WaitForGantrySafe_T1 := #s120_WaitForGantrySafe AND NOT #sStWtResetRel AND #sSst AND #iLoadGantrySafe;
END_REGION

REGION Network 40: STATE Num:120 Wait For Gantry Safe
   RUNG wire#powerrail
      Contact( #s120_WaitForGantrySafe )
      wire#w1
      I_Contact( #sStWtResetRel )
      I_Contact( #s120_WaitForGantrySafe_T1 )
      wire#w2
      Coil( #s120_WaitForGantrySafe )
   END_RUNG
   RUNG wire#powerrail
      Contact( #s100_WaitForOperatorDecision_T1 )
   END_RUNG wire#w1
   RUNG wire#powerrail
      Contact( #s90_ConfirmPartLoad_T2 )
   END_RUNG wire#w1
   RUNG wire#w2
      { S7_GenerateENO := "TRUE" } Move(in := 120, out1 => #StateNo)
   END_RUNG
   // the same network as SCL:
   #s120_WaitForGantrySafe := (#s120_WaitForGantrySafe OR #s100_WaitForOperatorDecision_T1 OR #s90_ConfirmPartLoad_T2) AND NOT #sStWtResetRel AND NOT #s120_WaitForGantrySafe_T1;
   IF #s120_WaitForGantrySafe THEN #StateNo := 120; END_IF;
END_REGION

REGION Network 41: Condition1 for STATE Num:121 Wait For RFID Write Over
   RUNG wire#powerrail
      Contact( #iRFWriteError )
      Coil( #c121_WaitForRFIDWriteOver_T1 )
   END_RUNG
   // the same network as SCL:
   #c121_WaitForRFIDWriteOver_T1 := #iRFWriteError;
END_REGION

REGION Network 42: Condition2 for STATE Num:121 Wait For RFID Write Over
   RUNG wire#powerrail
      Contact( #iRFWriteDone )
      Coil( #c121_WaitForRFIDWriteOver_T2 )
   END_RUNG
   // the same network as SCL:
   #c121_WaitForRFIDWriteOver_T2 := #iRFWriteDone;
END_REGION

REGION Network 43: Transition for STATE Num:121 Wait For RFID Write Over
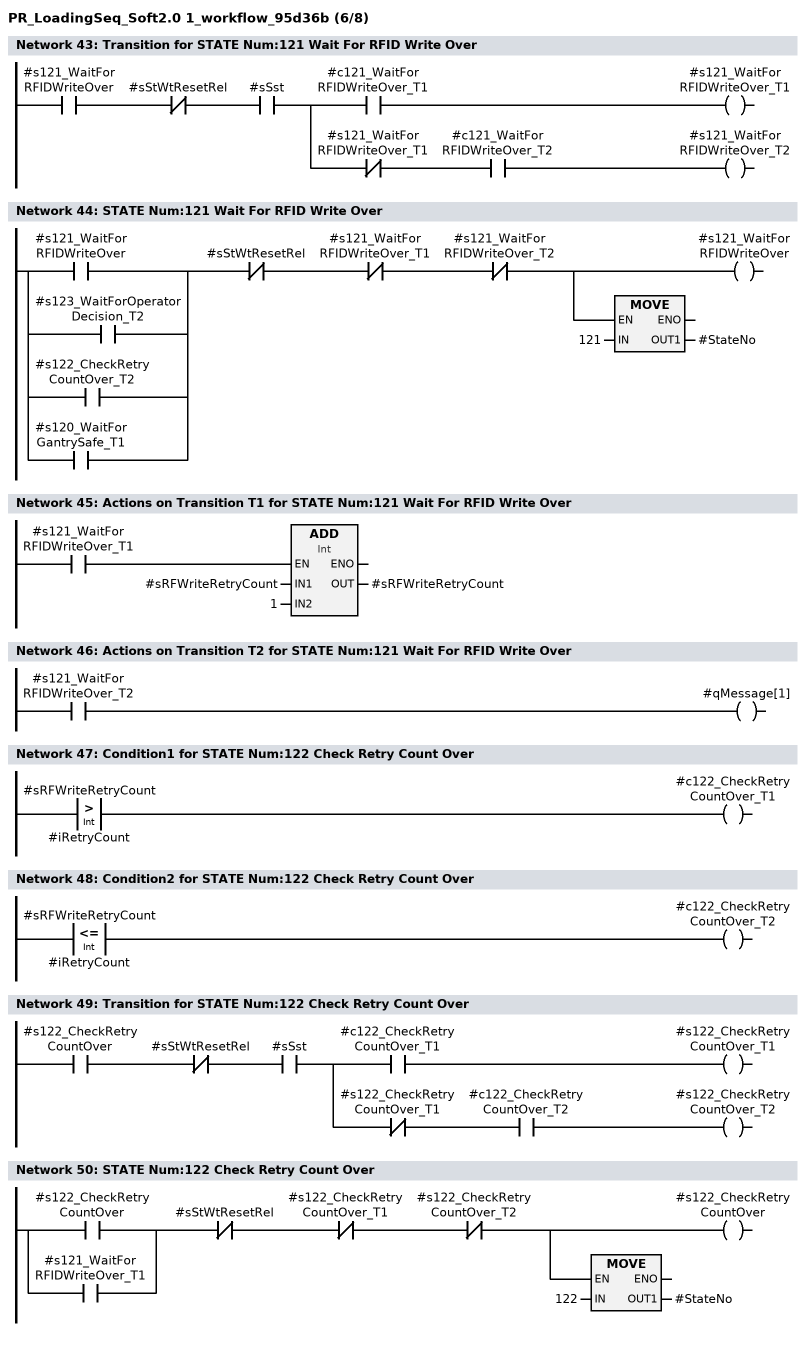
   RUNG wire#powerrail
      Contact( #s121_WaitForRFIDWriteOver )
      I_Contact( #sStWtResetRel )
      Contact( #sSst )
      wire#w1
      Contact( #c121_WaitForRFIDWriteOver_T1 )
      Coil( #s121_WaitForRFIDWriteOver_T1 )
   END_RUNG
   RUNG wire#w1
      I_Contact( #s121_WaitForRFIDWriteOver_T1 )
      Contact( #c121_WaitForRFIDWriteOver_T2 )
      Coil( #s121_WaitForRFIDWriteOver_T2 )
   END_RUNG
   // the same network as SCL:
   #_w1 := #s121_WaitForRFIDWriteOver AND NOT #sStWtResetRel AND #sSst;
   #s121_WaitForRFIDWriteOver_T1 := #_w1 AND #c121_WaitForRFIDWriteOver_T1;
   #s121_WaitForRFIDWriteOver_T2 := #_w1 AND NOT #s121_WaitForRFIDWriteOver_T1 AND #c121_WaitForRFIDWriteOver_T2;
END_REGION

REGION Network 44: STATE Num:121 Wait For RFID Write Over
   RUNG wire#powerrail
      Contact( #s121_WaitForRFIDWriteOver )
      wire#w1
      I_Contact( #sStWtResetRel )
      I_Contact( #s121_WaitForRFIDWriteOver_T1 )
      I_Contact( #s121_WaitForRFIDWriteOver_T2 )
      wire#w2
      Coil( #s121_WaitForRFIDWriteOver )
   END_RUNG
   RUNG wire#powerrail
      Contact( #s123_WaitForOperatorDecision_T2 )
   END_RUNG wire#w1
   RUNG wire#powerrail
      Contact( #s122_CheckRetryCountOver_T2 )
   END_RUNG wire#w1
   RUNG wire#powerrail
      Contact( #s120_WaitForGantrySafe_T1 )
   END_RUNG wire#w1
   RUNG wire#w2
      { S7_GenerateENO := "TRUE" } Move(in := 121, out1 => #StateNo)
   END_RUNG
   // the same network as SCL:
   #s121_WaitForRFIDWriteOver := (#s121_WaitForRFIDWriteOver OR #s123_WaitForOperatorDecision_T2 OR #s122_CheckRetryCountOver_T2 OR #s120_WaitForGantrySafe_T1) AND NOT #sStWtResetRel AND NOT #s121_WaitForRFIDWriteOver_T1 AND NOT #s121_WaitForRFIDWriteOver_T2;
   IF #s121_WaitForRFIDWriteOver THEN #StateNo := 121; END_IF;
END_REGION

REGION Network 45: Actions on Transition T1 for STATE Num:121 Wait For RFID Write Over
   RUNG wire#powerrail
      Contact( #s121_WaitForRFIDWriteOver_T1 )
      { S7_Templates := "SrcType := Int"; S7_GenerateENO := "TRUE" } Add(in1 := #sRFWriteRetryCount, in2 := 1, out => #sRFWriteRetryCount)
   END_RUNG
   // the same network as SCL:
   IF #s121_WaitForRFIDWriteOver_T1 THEN #sRFWriteRetryCount := #sRFWriteRetryCount + 1; END_IF;
END_REGION

REGION Network 46: Actions on Transition T2 for STATE Num:121 Wait For RFID Write Over
   RUNG wire#powerrail
      Contact( #s121_WaitForRFIDWriteOver_T2 )
      Coil( #qMessage[1] )
   END_RUNG
   // the same network as SCL:
   #qMessage[1] := #s121_WaitForRFIDWriteOver_T2;
END_REGION

REGION Network 47: Condition1 for STATE Num:122 Check Retry Count Over
   RUNG wire#powerrail
      { S7_Templates := "SrcType := Int" } GT_Contact(in1 := #sRFWriteRetryCount, in2 := #iRetryCount)
      Coil( #c122_CheckRetryCountOver_T1 )
   END_RUNG
   // the same network as SCL:
   #c122_CheckRetryCountOver_T1 := #sRFWriteRetryCount > #iRetryCount;
END_REGION

REGION Network 48: Condition2 for STATE Num:122 Check Retry Count Over
   RUNG wire#powerrail
      { S7_Templates := "SrcType := Int" } LE_Contact(in1 := #sRFWriteRetryCount, in2 := #iRetryCount)
      Coil( #c122_CheckRetryCountOver_T2 )
   END_RUNG
   // the same network as SCL:
   #c122_CheckRetryCountOver_T2 := #sRFWriteRetryCount <= #iRetryCount;
END_REGION

REGION Network 49: Transition for STATE Num:122 Check Retry Count Over
   RUNG wire#powerrail
      Contact( #s122_CheckRetryCountOver )
      I_Contact( #sStWtResetRel )
      Contact( #sSst )
      wire#w1
      Contact( #c122_CheckRetryCountOver_T1 )
      Coil( #s122_CheckRetryCountOver_T1 )
   END_RUNG
   RUNG wire#w1
      I_Contact( #s122_CheckRetryCountOver_T1 )
      Contact( #c122_CheckRetryCountOver_T2 )
      Coil( #s122_CheckRetryCountOver_T2 )
   END_RUNG
   // the same network as SCL:
   #_w1 := #s122_CheckRetryCountOver AND NOT #sStWtResetRel AND #sSst;
   #s122_CheckRetryCountOver_T1 := #_w1 AND #c122_CheckRetryCountOver_T1;
   #s122_CheckRetryCountOver_T2 := #_w1 AND NOT #s122_CheckRetryCountOver_T1 AND #c122_CheckRetryCountOver_T2;
END_REGION

REGION Network 50: STATE Num:122 Check Retry Count Over
   RUNG wire#powerrail
      Contact( #s122_CheckRetryCountOver )
      wire#w1
      I_Contact( #sStWtResetRel )
      I_Contact( #s122_CheckRetryCountOver_T1 )
      I_Contact( #s122_CheckRetryCountOver_T2 )
      wire#w2
      Coil( #s122_CheckRetryCountOver )
   END_RUNG
   RUNG wire#powerrail
      Contact( #s121_WaitForRFIDWriteOver_T1 )
   END_RUNG wire#w1
   RUNG wire#w2
      { S7_GenerateENO := "TRUE" } Move(in := 122, out1 => #StateNo)
   END_RUNG
   // the same network as SCL:
   #s122_CheckRetryCountOver := (#s122_CheckRetryCountOver OR #s121_WaitForRFIDWriteOver_T1) AND NOT #sStWtResetRel AND NOT #s122_CheckRetryCountOver_T1 AND NOT #s122_CheckRetryCountOver_T2;
   IF #s122_CheckRetryCountOver THEN #StateNo := 122; END_IF;
END_REGION

REGION Network 51: Actions on Transition T1 for STATE Num:122 Check Retry Count Over
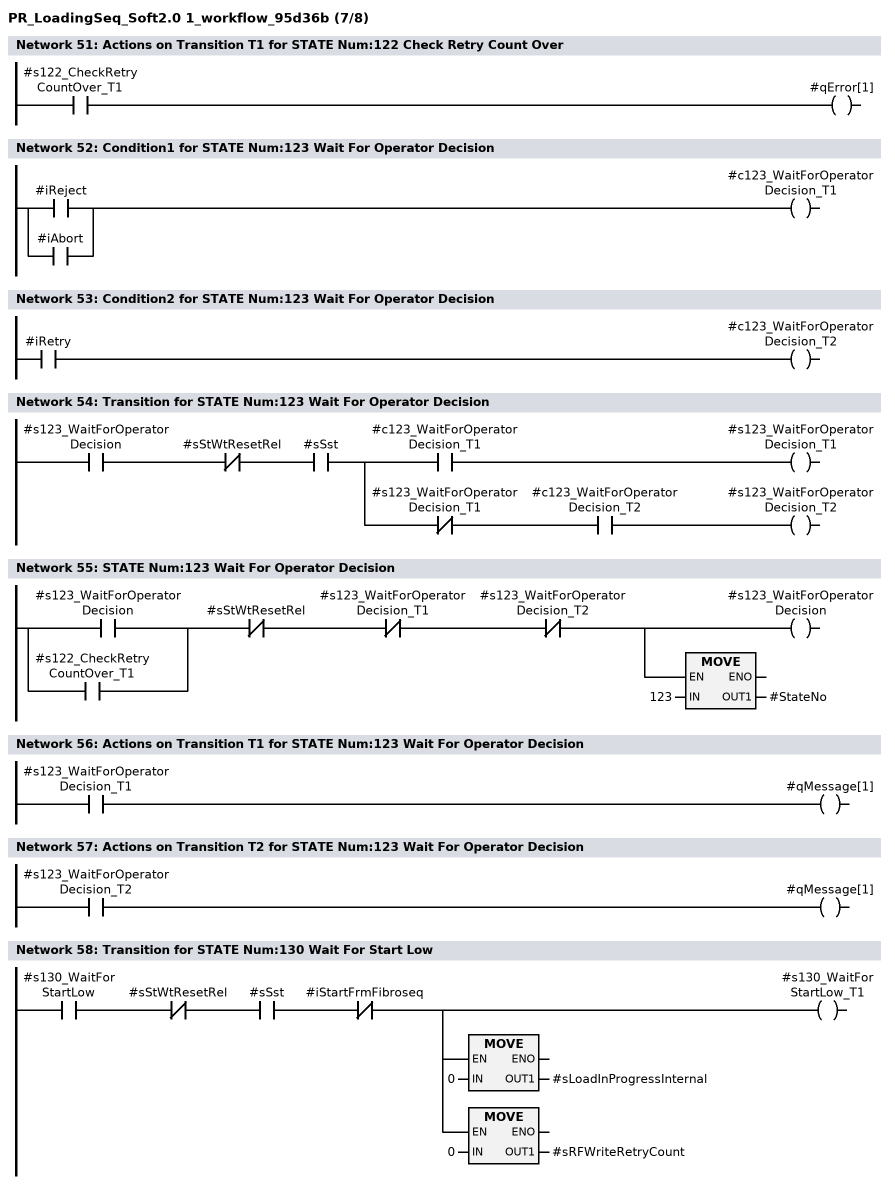
   RUNG wire#powerrail
      Contact( #s122_CheckRetryCountOver_T1 )
      Coil( #qError[1] )
   END_RUNG
   // the same network as SCL:
   #qError[1] := #s122_CheckRetryCountOver_T1;
END_REGION

REGION Network 52: Condition1 for STATE Num:123 Wait For Operator Decision
   RUNG wire#powerrail
      Contact( #iReject )
      wire#w1
      Coil( #c123_WaitForOperatorDecision_T1 )
   END_RUNG
   RUNG wire#powerrail
      Contact( #iAbort )
   END_RUNG wire#w1
   // the same network as SCL:
   #c123_WaitForOperatorDecision_T1 := #iReject OR #iAbort;
END_REGION

REGION Network 53: Condition2 for STATE Num:123 Wait For Operator Decision
   RUNG wire#powerrail
      Contact( #iRetry )
      Coil( #c123_WaitForOperatorDecision_T2 )
   END_RUNG
   // the same network as SCL:
   #c123_WaitForOperatorDecision_T2 := #iRetry;
END_REGION

REGION Network 54: Transition for STATE Num:123 Wait For Operator Decision
   RUNG wire#powerrail
      Contact( #s123_WaitForOperatorDecision )
      I_Contact( #sStWtResetRel )
      Contact( #sSst )
      wire#w1
      Contact( #c123_WaitForOperatorDecision_T1 )
      Coil( #s123_WaitForOperatorDecision_T1 )
   END_RUNG
   RUNG wire#w1
      I_Contact( #s123_WaitForOperatorDecision_T1 )
      Contact( #c123_WaitForOperatorDecision_T2 )
      Coil( #s123_WaitForOperatorDecision_T2 )
   END_RUNG
   // the same network as SCL:
   #_w1 := #s123_WaitForOperatorDecision AND NOT #sStWtResetRel AND #sSst;
   #s123_WaitForOperatorDecision_T1 := #_w1 AND #c123_WaitForOperatorDecision_T1;
   #s123_WaitForOperatorDecision_T2 := #_w1 AND NOT #s123_WaitForOperatorDecision_T1 AND #c123_WaitForOperatorDecision_T2;
END_REGION

REGION Network 55: STATE Num:123 Wait For Operator Decision
   RUNG wire#powerrail
      Contact( #s123_WaitForOperatorDecision )
      wire#w1
      I_Contact( #sStWtResetRel )
      I_Contact( #s123_WaitForOperatorDecision_T1 )
      I_Contact( #s123_WaitForOperatorDecision_T2 )
      wire#w2
      Coil( #s123_WaitForOperatorDecision )
   END_RUNG
   RUNG wire#powerrail
      Contact( #s122_CheckRetryCountOver_T1 )
   END_RUNG wire#w1
   RUNG wire#w2
      { S7_GenerateENO := "TRUE" } Move(in := 123, out1 => #StateNo)
   END_RUNG
   // the same network as SCL:
   #s123_WaitForOperatorDecision := (#s123_WaitForOperatorDecision OR #s122_CheckRetryCountOver_T1) AND NOT #sStWtResetRel AND NOT #s123_WaitForOperatorDecision_T1 AND NOT #s123_WaitForOperatorDecision_T2;
   IF #s123_WaitForOperatorDecision THEN #StateNo := 123; END_IF;
END_REGION

REGION Network 56: Actions on Transition T1 for STATE Num:123 Wait For Operator Decision
   RUNG wire#powerrail
      Contact( #s123_WaitForOperatorDecision_T1 )
      Coil( #qMessage[1] )
   END_RUNG
   // the same network as SCL:
   #qMessage[1] := #s123_WaitForOperatorDecision_T1;
END_REGION

REGION Network 57: Actions on Transition T2 for STATE Num:123 Wait For Operator Decision
   RUNG wire#powerrail
      Contact( #s123_WaitForOperatorDecision_T2 )
      Coil( #qMessage[1] )
   END_RUNG
   // the same network as SCL:
   #qMessage[1] := #s123_WaitForOperatorDecision_T2;
END_REGION

REGION Network 58: Transition for STATE Num:130 Wait For Start Low
   RUNG wire#powerrail
      Contact( #s130_WaitForStartLow )
      I_Contact( #sStWtResetRel )
      Contact( #sSst )
      I_Contact( #iStartFrmFibroseq )
      wire#w1
      Coil( #s130_WaitForStartLow_T1 )
   END_RUNG
   RUNG wire#w1
      Move(in := 0, out1 => #sLoadInProgressInternal)
   END_RUNG
   RUNG wire#w1
      Move(in := 0, out1 => #sRFWriteRetryCount)
   END_RUNG
   // the same network as SCL:
   #s130_WaitForStartLow_T1 := #s130_WaitForStartLow AND NOT #sStWtResetRel AND #sSst AND NOT #iStartFrmFibroseq;
   IF #s130_WaitForStartLow_T1 THEN
       #sLoadInProgressInternal := 0;
       #sRFWriteRetryCount := 0;
   END_IF;
END_REGION

REGION Network 59: STATE Num:130 Wait For Start Low
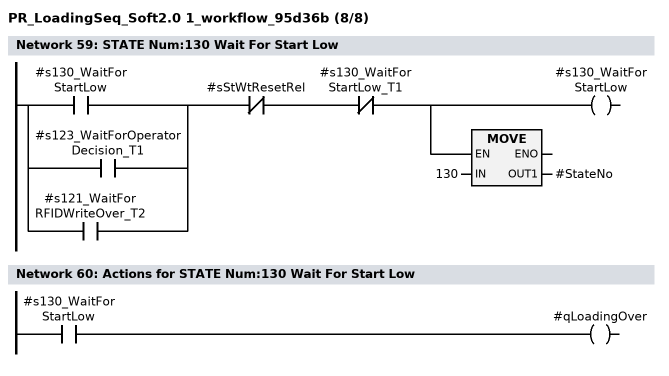
   RUNG wire#powerrail
      Contact( #s130_WaitForStartLow )
      wire#w1
      I_Contact( #sStWtResetRel )
      I_Contact( #s130_WaitForStartLow_T1 )
      wire#w2
      Coil( #s130_WaitForStartLow )
   END_RUNG
   RUNG wire#powerrail
      Contact( #s123_WaitForOperatorDecision_T1 )
   END_RUNG wire#w1
   RUNG wire#powerrail
      Contact( #s121_WaitForRFIDWriteOver_T2 )
   END_RUNG wire#w1
   RUNG wire#w2
      { S7_GenerateENO := "TRUE" } Move(in := 130, out1 => #StateNo)
   END_RUNG
   // the same network as SCL:
   #s130_WaitForStartLow := (#s130_WaitForStartLow OR #s123_WaitForOperatorDecision_T1 OR #s121_WaitForRFIDWriteOver_T2) AND NOT #sStWtResetRel AND NOT #s130_WaitForStartLow_T1;
   IF #s130_WaitForStartLow THEN #StateNo := 130; END_IF;
END_REGION

REGION Network 60: Actions for STATE Num:130 Wait For Start Low
   RUNG wire#powerrail
      Contact( #s130_WaitForStartLow )
      Coil( #qLoadingOver )
   END_RUNG
   // the same network as SCL:
   #qLoadingOver := #s130_WaitForStartLow;
END_REGION
END_FUNCTION_BLOCK
